FUNCTION maximum : LREAL
VAR_INPUT
	x: ARRAY[0..2] OF LREAL;
END_VAR
VAR
END_VAR


maximum := x[0];

IF x[0] < x[1] THEN 
    maximum := x[1];
END_IF;


IF maximum < x[2] THEN 
    maximum := x[2];
END_IF;

END_FUNCTION

(* stored: Version 1.1.0.1, ProductVersion 3.1.4024.9
   POU maximum: Id {b4de15a6-019e-4820-9ae4-4f8862d9701a}, SpecialFunc None *)
